(*
SPDX-FileCopyrightText: © 2026 Oleksandr Tiutyk <trofimich@gmail.com>
SPDX-License-Identifier: MIT
License: https://opensource.org/license/mit
*)

(*!
<summary>Represents an exception raised when an invalid workflow state transition is requested or attempted.</summary>
<description>
Dynamic copies are explicitly registered by Clone after construction; plain __NEW does not transfer ownership
to the task manager.
</description>
*)

{attribute 'enable_dynamic_creation'}
{attribute 'no_explicit_call' := 'do not call this function block directly'}
FUNCTION_BLOCK InvalidWorkflowTransitionException EXTENDS TOF_Core.GeneralException
	IMPLEMENTS IInvalidWorkflowTransitionException
VAR_STAT
	{attribute 'hide'} 
	_ClassName : STRING := __POUNAME();
END_VAR

(*!
<summary>Borrows the initialized class name used in diagnostics.</summary>
<description>
Returns initialized metadata storage without allocation. Callers must not modify the returned string.
Derived function blocks must use distinct initialized static storage when overriding this metadata.
</description>
*)
{attribute 'monitoring' := 'call'}
PROPERTY ClassName : REFERENCE TO STRING
GET
ClassName REF= _ClassName;
END_GET
END_PROPERTY

(*!
<summary>Creates a task-owned copy of this exception and its diagnostic payload.</summary>
<description>
Registers the newly constructed instance before copying payload, outside FB_init. Registration failure
releases the unregistered instance and raises a terminal error; copy failure leaves the registered instance
owned by the task manager for cleanup. Custom overrides must follow the same ownership sequence. The returned
reference is borrowed until task cleanup and must not be deleted by the caller.
</description>
*)
METHOD Clone : TOF_Core.IObject
VAR
	exceptionClone : POINTER TO InvalidWorkflowTransitionException;
END_VAR
exceptionClone := __NEW(InvalidWorkflowTransitionException);

IF exceptionClone = 0 THEN
	TOF_Core.DynamicMemoryManager.RaiseAllocationFailure();
END_IF

TOF_Core.DynamicMemoryManager.RegisterAutoDisposedObject(autoDisposedObject := exceptionClone^);

exceptionClone^.CopyGeneralFields(sourceException := THIS^);

Clone := exceptionClone^;
END_METHOD

(*!
<summary>Borrows the compiler-initialized library namespace.</summary>
<description>
Borrows storage from the live internal namespace provider. Reacquire references after application
reinitialization or relocation. Treat the reference as read-only; no ownership or synchronization is provided.
</description>
*)
{attribute 'monitoring' := 'call'}
PROPERTY NamespaceName : REFERENCE TO STRING
GET
NamespaceName REF= CurrentNamespace.Name;
END_GET
END_PROPERTY

(*!
<summary>Reports the size of this concrete function block instance in bytes.</summary>
<description>
Reports the instance layout rather than dynamic allocations owned by its fields. A derived function block
with a different layout must override this property; the value does not grant disposal rights.
</description>
*)
{attribute 'monitoring' := 'call'}
PROPERTY SelfSize : ULINT
GET
SelfSize := XSIZEOF(THIS^);
END_GET
END_PROPERTY

(*!
<summary>Formats the invalid state transition diagnostic and raises this exception.</summary>
<description>
Formats the diagnostic without heap allocation during message preparation and propagates the exception.
</description>
<param name="sourceNamespaceName">Namespace of the POU raising the exception.</param>
<param name="sourceClassName">Class name of the workflow element where the transition was rejected.</param>
<param name="sourcePOUName">Method or property name where the transition was attempted.</param>
<param name="sourcePosition">Source position identifier.</param>
<param name="fromState">Current state of the workflow element.</param>
<param name="toState">Rejected target state.</param>
*)
METHOD Throw
VAR_INPUT
	sourceNamespaceName : STRING;
	sourceClassName : STRING;
	sourcePOUName : STRING;
	sourcePosition : STRING;
	fromState : WORKFLOW_ELEMENT_STATE;
	toState : WORKFLOW_ELEMENT_STATE;
END_VAR
VAR
	message : TOF_Core.ERROR_MESSAGE;
END_VAR
message := TOF_Core.WideStrings.Concat255(
	"Transition from state '",
	TO_WSTRING(fromState),
	"' to state '",
	TO_WSTRING(toState),
	"' is not allowed");

InternalThrow(
	sourceNamespaceName := sourceNamespaceName,
	sourceClassName := sourceClassName,
	sourcePOUName := sourcePOUName,
	sourcePosition := sourcePosition,
	message := message,
	errorCode := 0,
	innerException := 0
);
END_METHOD

END_FUNCTION_BLOCK

(* stored: Version 1.1.0.1
   POU InvalidWorkflowTransitionException: Id {4f38afb5-d1df-4cda-9265-546e40bc6542}, SpecialFunc None
   Property ClassName: Id {2344dbe6-d582-4933-b2fa-6b01450c7cc8}
   Get Get: Id {913a6212-cfb0-489c-86ff-34ac85c54435}
   Method Clone: Id {e5a7d856-90d1-4514-a381-acaaf01ec409}
   Property NamespaceName: Id {34567feb-3e62-4418-9e99-7e3be338908d}
   Get Get: Id {962acf80-b1e1-44e0-8ae4-6f8ce61ac7db}
   Property SelfSize: Id {6e91bb6e-b109-459e-ad7c-7b9bfdf49e97}
   Get Get: Id {2475efcb-21ff-4c76-9a35-80543d39595c}
   Method Throw: Id {06f59df7-586a-4456-b537-5f6e9d8adcc7} *)
